(* IEC 61131-3 sources: plc-st-coding-agent/progress/evidence/f14_v3_parallel_20261112/jobs/codex_deepseek-v4pro (part 2) *)

(* ---- public-medium-05.candidate_02.st ---- *)
FUNCTION_BLOCK AutomatedProductionLine
VAR_INPUT
    Mode : BOOL;
    ForwardButton : BOOL;
    ReverseButton : BOOL;
    SensorA : BOOL;
    SensorB : BOOL;
    SensorC : BOOL;
    ButtonA : BOOL;
    ButtonB : BOOL;
    ButtonC : BOOL;
END_VAR
VAR_OUTPUT
    MotorForward : BOOL;
    MotorReverse : BOOL;
    CompletionLight : BOOL;
END_VAR
VAR
    SequenceStep : INT := 0;
END_VAR

MotorForward := FALSE;
MotorReverse := FALSE;
CompletionLight := FALSE;

IF NOT Mode THEN
    MotorForward := ForwardButton AND NOT ReverseButton;
    MotorReverse := ReverseButton AND NOT ForwardButton;
ELSE
    MotorReverse := FALSE;

    CASE SequenceStep OF
        0:
            IF SensorA AND ButtonA THEN
                SequenceStep := 1;
            END_IF;

        1:
            MotorForward := TRUE;
            IF SensorB THEN
                MotorForward := FALSE;
                SequenceStep := 2;
            END_IF;

        2:
            IF ButtonB THEN
                SequenceStep := 3;
            END_IF;

        3:
            MotorForward := TRUE;
            IF SensorC THEN
                MotorForward := FALSE;
                SequenceStep := 4;
            END_IF;

        4:
            IF ButtonC THEN
                SequenceStep := 5;
            END_IF;

        5:
            CompletionLight := SensorC;
            IF NOT SensorC THEN
                CompletionLight := FALSE;
                SequenceStep := 0;
            END_IF;
    END_CASE;
END_IF;

END_FUNCTION_BLOCK

(* ---- public-medium-05.raw_candidate_01.st ---- *)
FUNCTION_BLOCK AutomatedProductionLine
VAR
    SequenceStep : INT := 0;
END_VAR

MotorForward := FALSE;
MotorReverse := FALSE;
CompletionLight := FALSE;

IF NOT Mode THEN
    MotorForward := ForwardButton AND NOT ReverseButton;
    MotorReverse := ReverseButton AND NOT ForwardButton;
    CompletionLight := FALSE;
ELSE
    MotorReverse := FALSE;

    CASE SequenceStep OF
        0:
            IF SensorA AND ButtonA THEN
                SequenceStep := 1;
            END_IF;

        1:
            MotorForward := TRUE;
            IF SensorB THEN
                MotorForward := FALSE;
                SequenceStep := 2;
            END_IF;

        2:
            IF ButtonB THEN
                SequenceStep := 3;
            END_IF;

        3:
            MotorForward := TRUE;
            IF SensorC THEN
                MotorForward := FALSE;
                SequenceStep := 4;
            END_IF;

        4:
            IF ButtonC THEN
                SequenceStep := 5;
            END_IF;

        5:
            CompletionLight := SensorC;
            IF NOT SensorC THEN
                CompletionLight := FALSE;
                SequenceStep := 0;
            END_IF;
    END_CASE;
END_IF;

END_FUNCTION_BLOCK

(* ---- public-medium-05.raw_candidate_02.st ---- *)
FUNCTION_BLOCK AutomatedProductionLine
VAR_INPUT
    Mode : BOOL;
    ForwardButton : BOOL;
    ReverseButton : BOOL;
    SensorA : BOOL;
    SensorB : BOOL;
    SensorC : BOOL;
    ButtonA : BOOL;
    ButtonB : BOOL;
    ButtonC : BOOL;
END_VAR
VAR_OUTPUT
    MotorForward : BOOL;
    MotorReverse : BOOL;
    CompletionLight : BOOL;
END_VAR
VAR
    SequenceStep : INT := 0;
END_VAR

MotorForward := FALSE;
MotorReverse := FALSE;
CompletionLight := FALSE;

IF NOT Mode THEN
    MotorForward := ForwardButton AND NOT ReverseButton;
    MotorReverse := ReverseButton AND NOT ForwardButton;
ELSE
    MotorReverse := FALSE;

    CASE SequenceStep OF
        0:
            IF SensorA AND ButtonA THEN
                SequenceStep := 1;
            END_IF;

        1:
            MotorForward := TRUE;
            IF SensorB THEN
                MotorForward := FALSE;
                SequenceStep := 2;
            END_IF;

        2:
            IF ButtonB THEN
                SequenceStep := 3;
            END_IF;

        3:
            MotorForward := TRUE;
            IF SensorC THEN
                MotorForward := FALSE;
                SequenceStep := 4;
            END_IF;

        4:
            IF ButtonC THEN
                SequenceStep := 5;
            END_IF;

        5:
            CompletionLight := SensorC;
            IF NOT SensorC THEN
                CompletionLight := FALSE;
                SequenceStep := 0;
            END_IF;
    END_CASE;
END_IF;

END_FUNCTION_BLOCK

(* ---- public-medium-06.candidate_01.st ---- *)
FUNCTION_BLOCK SlabThicknessAlarmFaultHistory
VAR_INPUT
    THICKNESS_FAULT : BOOL;
    THICKNESS_SIGNAL_VALID : BOOL;
    CUTTING_RUN : BOOL;
    FaultTimestamp : DINT;
    CycleTime : TIME;
END_VAR
VAR_OUTPUT
    THICKNESS_ALARM : BOOL;
    Slab_Fault_Counter : UINT;
    Slab_Runtime_Accumulator : LTIME;
    Slab_Fault_History : ARRAY[0..4] OF DINT;
END_VAR
VAR
    Initialized : BOOL := FALSE;
    CurrentValidFault : BOOL;
    LastValidFault : BOOL := FALSE;
    AlarmHolding : BOOL := FALSE;
    AlarmHoldTimer : TIME := T#0ms;
    ArrayIndex : INT;
END_VAR

IF NOT Initialized THEN
    THICKNESS_ALARM := FALSE;
    Slab_Fault_Counter := 0;
    Slab_Runtime_Accumulator := TIME_TO_LTIME(T#0ms);
    FOR ArrayIndex := 0 TO 4 DO
        Slab_Fault_History[ArrayIndex] := 0;
    END_FOR;
    AlarmHolding := FALSE;
    AlarmHoldTimer := T#0ms;
    LastValidFault := THICKNESS_SIGNAL_VALID AND THICKNESS_FAULT;
    Initialized := TRUE;
END_IF;

IF NOT THICKNESS_SIGNAL_VALID THEN
    THICKNESS_ALARM := FALSE;
    AlarmHolding := FALSE;
    AlarmHoldTimer := T#0ms;
    LastValidFault := FALSE;
ELSE
    CurrentValidFault := THICKNESS_FAULT;

    IF CurrentValidFault AND NOT LastValidFault THEN
        Slab_Fault_Counter := Slab_Fault_Counter + 1;
        FOR ArrayIndex := 4 TO 1 BY -1 DO
            Slab_Fault_History[ArrayIndex] := Slab_Fault_History[ArrayIndex - 1];
        END_FOR;
        Slab_Fault_History[0] := FaultTimestamp;
    END_IF;

    IF CurrentValidFault THEN
        THICKNESS_ALARM := TRUE;
        AlarmHolding := TRUE;
        AlarmHoldTimer := T#0ms;
    ELSIF AlarmHolding THEN
        AlarmHoldTimer := AlarmHoldTimer + CycleTime;
        THICKNESS_ALARM := TRUE;
        IF AlarmHoldTimer >= T#500ms THEN
            THICKNESS_ALARM := FALSE;
            AlarmHolding := FALSE;
            AlarmHoldTimer := T#0ms;
        END_IF;
    ELSE
        THICKNESS_ALARM := FALSE;
    END_IF;

    LastValidFault := CurrentValidFault;
END_IF;

IF CUTTING_RUN AND THICKNESS_SIGNAL_VALID AND NOT THICKNESS_FAULT THEN
    Slab_Runtime_Accumulator := Slab_Runtime_Accumulator + TIME_TO_LTIME(CycleTime);
END_IF;

END_FUNCTION_BLOCK

(* ---- public-medium-06.candidate_02.st ---- *)
FUNCTION_BLOCK SlabThicknessAlarmFaultHistory
VAR_INPUT
    THICKNESS_FAULT : BOOL;
    THICKNESS_SIGNAL_VALID : BOOL;
    CUTTING_RUN : BOOL;
    FaultTimestamp : DINT;
    CycleTime : TIME;
END_VAR
VAR_OUTPUT
    THICKNESS_ALARM : BOOL;
    Slab_Fault_Counter : UINT;
    Slab_Runtime_Accumulator : LTIME;
    Slab_Fault_History : ARRAY[0..4] OF DINT;
END_VAR
VAR
    PowerUp : BOOL := TRUE;
    LastValidFault : BOOL := FALSE;
    CurrentFault : BOOL;
    AlarmHoldActive : BOOL := FALSE;
    AlarmHoldElapsed : TIME := T#0ms;
    LoopIndex : INT;
END_VAR

IF PowerUp THEN
    THICKNESS_ALARM := FALSE;
    Slab_Fault_Counter := 0;
    Slab_Runtime_Accumulator := TIME_TO_LTIME(T#0ms);
    FOR LoopIndex := 0 TO 4 DO
        Slab_Fault_History[LoopIndex] := 0;
    END_FOR;
    LastValidFault := FALSE;
    AlarmHoldActive := FALSE;
    AlarmHoldElapsed := T#0ms;
    PowerUp := FALSE;
END_IF;

IF NOT THICKNESS_SIGNAL_VALID THEN
    THICKNESS_ALARM := FALSE;
    AlarmHoldActive := FALSE;
    AlarmHoldElapsed := T#0ms;
    LastValidFault := FALSE;
ELSE
    CurrentFault := THICKNESS_FAULT;

    IF CurrentFault AND NOT LastValidFault THEN
        Slab_Fault_Counter := Slab_Fault_Counter + 1;
        FOR LoopIndex := 4 TO 1 BY -1 DO
            Slab_Fault_History[LoopIndex] := Slab_Fault_History[LoopIndex - 1];
        END_FOR;
        Slab_Fault_History[0] := FaultTimestamp;
    END_IF;

    IF CurrentFault THEN
        THICKNESS_ALARM := TRUE;
        AlarmHoldActive := TRUE;
        AlarmHoldElapsed := T#0ms;
    ELSIF AlarmHoldActive THEN
        AlarmHoldElapsed := AlarmHoldElapsed + CycleTime;
        IF AlarmHoldElapsed >= T#500ms THEN
            THICKNESS_ALARM := FALSE;
            AlarmHoldActive := FALSE;
            AlarmHoldElapsed := T#0ms;
        ELSE
            THICKNESS_ALARM := TRUE;
        END_IF;
    ELSE
        THICKNESS_ALARM := FALSE;
    END_IF;

    LastValidFault := CurrentFault;
END_IF;

IF CUTTING_RUN AND THICKNESS_SIGNAL_VALID AND NOT THICKNESS_FAULT THEN
    Slab_Runtime_Accumulator := Slab_Runtime_Accumulator + TIME_TO_LTIME(CycleTime);
END_IF;

END_FUNCTION_BLOCK

(* ---- public-medium-06.raw_candidate_01.st ---- *)
FUNCTION_BLOCK SlabThicknessAlarmFaultHistory
VAR_INPUT
    THICKNESS_FAULT : BOOL;
    THICKNESS_SIGNAL_VALID : BOOL;
    CUTTING_RUN : BOOL;
    FaultTimestamp : DINT;
    CycleTime : TIME;
END_VAR
VAR_OUTPUT
    THICKNESS_ALARM : BOOL;
    Slab_Fault_Counter : UINT;
    Slab_Runtime_Accumulator : LTIME;
    Slab_Fault_History : ARRAY[0..4] OF DINT;
END_VAR
VAR
    Initialized : BOOL := FALSE;
    CurrentValidFault : BOOL;
    LastValidFault : BOOL := FALSE;
    AlarmHolding : BOOL := FALSE;
    AlarmHoldTimer : TIME := T#0ms;
    ArrayIndex : INT;
END_VAR

IF NOT Initialized THEN
    THICKNESS_ALARM := FALSE;
    Slab_Fault_Counter := 0;
    Slab_Runtime_Accumulator := TIME_TO_LTIME(T#0ms);
    FOR ArrayIndex := 0 TO 4 DO
        Slab_Fault_History[ArrayIndex] := 0;
    END_FOR;
    AlarmHolding := FALSE;
    AlarmHoldTimer := T#0ms;
    LastValidFault := THICKNESS_SIGNAL_VALID AND THICKNESS_FAULT;
    Initialized := TRUE;
END_IF;

IF NOT THICKNESS_SIGNAL_VALID THEN
    THICKNESS_ALARM := FALSE;
    AlarmHolding := FALSE;
    AlarmHoldTimer := T#0ms;
    LastValidFault := FALSE;
ELSE
    CurrentValidFault := THICKNESS_FAULT;

    IF CurrentValidFault AND NOT LastValidFault THEN
        Slab_Fault_Counter := Slab_Fault_Counter + 1;
        FOR ArrayIndex := 4 TO 1 BY -1 DO
            Slab_Fault_History[ArrayIndex] := Slab_Fault_History[ArrayIndex - 1];
        END_FOR;
        Slab_Fault_History[0] := FaultTimestamp;
    END_IF;

    IF CurrentValidFault THEN
        THICKNESS_ALARM := TRUE;
        AlarmHolding := TRUE;
        AlarmHoldTimer := T#0ms;
    ELSIF AlarmHolding THEN
        AlarmHoldTimer := AlarmHoldTimer + CycleTime;
        THICKNESS_ALARM := TRUE;
        IF AlarmHoldTimer >= T#500ms THEN
            THICKNESS_ALARM := FALSE;
            AlarmHolding := FALSE;
            AlarmHoldTimer := T#0ms;
        END_IF;
    ELSE
        THICKNESS_ALARM := FALSE;
    END_IF;

    LastValidFault := CurrentValidFault;
END_IF;

IF CUTTING_RUN AND THICKNESS_SIGNAL_VALID AND NOT THICKNESS_FAULT THEN
    Slab_Runtime_Accumulator := Slab_Runtime_Accumulator + TIME_TO_LTIME(CycleTime);
END_IF;

END_FUNCTION_BLOCK

(* ---- public-medium-06.raw_candidate_02.st ---- *)
FUNCTION_BLOCK SlabThicknessAlarmFaultHistory
VAR_INPUT
    THICKNESS_FAULT : BOOL;
    THICKNESS_SIGNAL_VALID : BOOL;
    CUTTING_RUN : BOOL;
    FaultTimestamp : DINT;
    CycleTime : TIME;
END_VAR
VAR_OUTPUT
    THICKNESS_ALARM : BOOL;
    Slab_Fault_Counter : UINT;
    Slab_Runtime_Accumulator : LTIME;
    Slab_Fault_History : ARRAY[0..4] OF DINT;
END_VAR
VAR
    PowerUp : BOOL := TRUE;
    LastValidFault : BOOL := FALSE;
    CurrentFault : BOOL;
    AlarmHoldActive : BOOL := FALSE;
    AlarmHoldElapsed : TIME := T#0ms;
    LoopIndex : INT;
END_VAR

IF PowerUp THEN
    THICKNESS_ALARM := FALSE;
    Slab_Fault_Counter := 0;
    Slab_Runtime_Accumulator := TIME_TO_LTIME(T#0ms);
    FOR LoopIndex := 0 TO 4 DO
        Slab_Fault_History[LoopIndex] := 0;
    END_FOR;
    LastValidFault := FALSE;
    AlarmHoldActive := FALSE;
    AlarmHoldElapsed := T#0ms;
    PowerUp := FALSE;
END_IF;

IF NOT THICKNESS_SIGNAL_VALID THEN
    THICKNESS_ALARM := FALSE;
    AlarmHoldActive := FALSE;
    AlarmHoldElapsed := T#0ms;
    LastValidFault := FALSE;
ELSE
    CurrentFault := THICKNESS_FAULT;

    IF CurrentFault AND NOT LastValidFault THEN
        Slab_Fault_Counter := Slab_Fault_Counter + 1;
        FOR LoopIndex := 4 TO 1 BY -1 DO
            Slab_Fault_History[LoopIndex] := Slab_Fault_History[LoopIndex - 1];
        END_FOR;
        Slab_Fault_History[0] := FaultTimestamp;
    END_IF;

    IF CurrentFault THEN
        THICKNESS_ALARM := TRUE;
        AlarmHoldActive := TRUE;
        AlarmHoldElapsed := T#0ms;
    ELSIF AlarmHoldActive THEN
        AlarmHoldElapsed := AlarmHoldElapsed + CycleTime;
        IF AlarmHoldElapsed >= T#500ms THEN
            THICKNESS_ALARM := FALSE;
            AlarmHoldActive := FALSE;
            AlarmHoldElapsed := T#0ms;
        ELSE
            THICKNESS_ALARM := TRUE;
        END_IF;
    ELSE
        THICKNESS_ALARM := FALSE;
    END_IF;

    LastValidFault := CurrentFault;
END_IF;

IF CUTTING_RUN AND THICKNESS_SIGNAL_VALID AND NOT THICKNESS_FAULT THEN
    Slab_Runtime_Accumulator := Slab_Runtime_Accumulator + TIME_TO_LTIME(CycleTime);
END_IF;

END_FUNCTION_BLOCK

(* ---- public-medium-07.candidate_01.st ---- *)
FUNCTION_BLOCK OfficeHVACMultiModeControl
VAR_INPUT
    OCCUPANCY_DETECTED : BOOL;
    ENERGY_SAVING_MODE : BOOL;
    HVAC_MODE_SELECTOR : INT;
END_VAR
VAR_OUTPUT
    SUPPLY_FAN_RUN : BOOL := FALSE;
    TEMP_SETPOINT_ADJUST : INT := 0;
END_VAR
VAR
    fan_timer : TON;
    setpoint_calc : INT;
END_VAR

fan_timer(IN := OCCUPANCY_DETECTED AND (HVAC_MODE_SELECTOR <> 3), PT := T#30S);
SUPPLY_FAN_RUN := fan_timer.Q;

CASE HVAC_MODE_SELECTOR OF
    0:
        IF OCCUPANCY_DETECTED THEN
            setpoint_calc := 0;
        ELSIF ENERGY_SAVING_MODE THEN
            setpoint_calc := 3;
        ELSE
            setpoint_calc := 2;
        END_IF;
    1:
        IF OCCUPANCY_DETECTED THEN
            setpoint_calc := 0;
        ELSE
            setpoint_calc := 1;
        END_IF;
    2:
        IF OCCUPANCY_DETECTED THEN
            setpoint_calc := 0;
        ELSE
            setpoint_calc := 4;
        END_IF;
    3:
        setpoint_calc := 4;
    ELSE
        setpoint_calc := 0;
END_CASE;

IF setpoint_calc > 4 THEN
    TEMP_SETPOINT_ADJUST := 4;
ELSIF setpoint_calc < -4 THEN
    TEMP_SETPOINT_ADJUST := -4;
ELSE
    TEMP_SETPOINT_ADJUST := setpoint_calc;
END_IF;
END_FUNCTION_BLOCK

(* ---- public-medium-07.raw_candidate_01.st ---- *)
FUNCTION_BLOCK OfficeHVACMultiModeControl
VAR_INPUT
    OCCUPANCY_DETECTED : BOOL;
    ENERGY_SAVING_MODE : BOOL;
    HVAC_MODE_SELECTOR : INT;
END_VAR
VAR_OUTPUT
    SUPPLY_FAN_RUN : BOOL := FALSE;
    TEMP_SETPOINT_ADJUST : INT := 0;
END_VAR
VAR
    fan_timer : TON;
    setpoint_calc : INT;
END_VAR

fan_timer(IN := OCCUPANCY_DETECTED AND (HVAC_MODE_SELECTOR <> 3), PT := T#30S);
SUPPLY_FAN_RUN := fan_timer.Q;

CASE HVAC_MODE_SELECTOR OF
    0:
        IF OCCUPANCY_DETECTED THEN
            setpoint_calc := 0;
        ELSIF ENERGY_SAVING_MODE THEN
            setpoint_calc := 3;
        ELSE
            setpoint_calc := 2;
        END_IF;
    1:
        IF OCCUPANCY_DETECTED THEN
            setpoint_calc := 0;
        ELSE
            setpoint_calc := 1;
        END_IF;
    2:
        IF OCCUPANCY_DETECTED THEN
            setpoint_calc := 0;
        ELSE
            setpoint_calc := 4;
        END_IF;
    3:
        setpoint_calc := 4;
    ELSE
        setpoint_calc := 0;
END_CASE;

IF setpoint_calc > 4 THEN
    TEMP_SETPOINT_ADJUST := 4;
ELSIF setpoint_calc < -4 THEN
    TEMP_SETPOINT_ADJUST := -4;
ELSE
    TEMP_SETPOINT_ADJUST := setpoint_calc;
END_IF;
END_FUNCTION_BLOCK

(* ---- public-medium-08.candidate_01.st ---- *)
FUNCTION_BLOCK IPv4Parser
VAR_INPUT
    ipText : STRING(254);
END_VAR
VAR_OUTPUT
    ipValue : UDINT;
END_VAR
VAR
    bValid : BOOL;
    iPos : INT;
    iLength : INT;
    iCharCode : INT;
    uiCurrentValue : UDINT;
    uiDigitCount : UDINT;
    uiCompletedSegments : UDINT;
    uiAddress : UDINT;
END_VAR

ipValue := 0;
uiAddress := 0;
uiCurrentValue := 0;
uiDigitCount := 0;
uiCompletedSegments := 0;
bValid := TRUE;
iLength := LEN(ipText);

IF (iLength > 0) AND (iLength <= 15) THEN
    FOR iPos := 1 TO iLength BY 1 DO
        iCharCode := BYTE_TO_INT(ipText[iPos]);

        IF (iCharCode >= 48) AND (iCharCode <= 57) THEN
            uiCurrentValue := uiCurrentValue * 10 + INT_TO_UDINT(iCharCode - 48);
            uiDigitCount := uiDigitCount + 1;

            IF uiCurrentValue > 255 THEN
                bValid := FALSE;
                EXIT;
            END_IF;

        ELSIF iCharCode = 46 THEN
            IF (uiDigitCount = 0) OR (uiCompletedSegments >= 3) THEN
                bValid := FALSE;
                EXIT;
            END_IF;

            uiAddress := uiAddress * 256 + uiCurrentValue;
            uiCompletedSegments := uiCompletedSegments + 1;
            uiCurrentValue := 0;
            uiDigitCount := 0;

        ELSE
            bValid := FALSE;
            EXIT;
        END_IF;
    END_FOR;
ELSE
    bValid := FALSE;
END_IF;

IF bValid THEN
    IF (uiDigitCount = 0) OR (uiCompletedSegments <> 3) THEN
        bValid := FALSE;
    ELSE
        uiAddress := uiAddress * 256 + uiCurrentValue;
        ipValue := uiAddress;
    END_IF;
END_IF;

END_FUNCTION_BLOCK

(* ---- public-medium-08.raw_candidate_01.st ---- *)
FUNCTION_BLOCK IPv4Parser
VAR_INPUT
    ipText : STRING(254);
END_VAR
VAR_OUTPUT
    ipValue : UDINT;
END_VAR
VAR
    bValid : BOOL;
    iPos : INT;
    iLength : INT;
    iCharCode : INT;
    uiCurrentValue : UDINT;
    uiDigitCount : UDINT;
    uiCompletedSegments : UDINT;
    uiAddress : UDINT;
END_VAR

ipValue := 0;
uiAddress := 0;
uiCurrentValue := 0;
uiDigitCount := 0;
uiCompletedSegments := 0;
bValid := TRUE;
iLength := LEN(ipText);

IF (iLength > 0) AND (iLength <= 15) THEN
    FOR iPos := 1 TO iLength BY 1 DO
        iCharCode := BYTE_TO_INT(ipText[iPos]);

        IF (iCharCode >= 48) AND (iCharCode <= 57) THEN
            uiCurrentValue := uiCurrentValue * 10 + INT_TO_UDINT(iCharCode - 48);
            uiDigitCount := uiDigitCount + 1;

            IF uiCurrentValue > 255 THEN
                bValid := FALSE;
                EXIT;
            END_IF;

        ELSIF iCharCode = 46 THEN
            IF (uiDigitCount = 0) OR (uiCompletedSegments >= 3) THEN
                bValid := FALSE;
                EXIT;
            END_IF;

            uiAddress := uiAddress * 256 + uiCurrentValue;
            uiCompletedSegments := uiCompletedSegments + 1;
            uiCurrentValue := 0;
            uiDigitCount := 0;

        ELSE
            bValid := FALSE;
            EXIT;
        END_IF;
    END_FOR;
ELSE
    bValid := FALSE;
END_IF;

IF bValid THEN
    IF (uiDigitCount = 0) OR (uiCompletedSegments <> 3) THEN
        bValid := FALSE;
    ELSE
        uiAddress := uiAddress * 256 + uiCurrentValue;
        ipValue := uiAddress;
    END_IF;
END_IF;

END_FUNCTION_BLOCK

(* ---- self-easy-01.candidate_01.st ---- *)
FUNCTION_BLOCK FB
VAR_INPUT
    enable : BOOL;
    values : ARRAY[1..8] OF INT;
    count : INT;
    avgEnable : BOOL;
END_VAR
VAR_OUTPUT
    avgOut : REAL;
END_VAR
VAR
    sampleCount : INT;
    total : LINT;
    idx : INT;
END_VAR

IF enable AND avgEnable AND (count > 0) THEN
    IF count > 8 THEN
        sampleCount := 8;
    ELSE
        sampleCount := count;
    END_IF;

    total := LINT#0;

    FOR idx := 1 TO sampleCount BY 1 DO
        total := total + INT_TO_LINT(values[idx]);
    END_FOR;

    avgOut := LINT_TO_REAL(total) / INT_TO_REAL(sampleCount);
END_IF;

END_FUNCTION_BLOCK

(* ---- self-easy-01.raw_candidate_01.st ---- *)
FUNCTION_BLOCK FB
VAR_INPUT
    enable : BOOL;
    values : ARRAY[1..8] OF INT;
    count : INT;
    avgEnable : BOOL;
END_VAR
VAR_OUTPUT
    avgOut : REAL;
END_VAR
VAR
    sampleCount : INT;
    total : LINT;
    idx : INT;
END_VAR

IF enable AND avgEnable AND (count > 0) THEN
    IF count > 8 THEN
        sampleCount := 8;
    ELSE
        sampleCount := count;
    END_IF;

    total := LINT#0;

    FOR idx := 1 TO sampleCount BY 1 DO
        total := total + INT_TO_LINT(values[idx]);
    END_FOR;

    avgOut := LINT_TO_REAL(total) / INT_TO_REAL(sampleCount);
END_IF;

END_FUNCTION_BLOCK

(* ---- self-easy-02.candidate_01.st ---- *)
FUNCTION_BLOCK FB
VAR_INPUT
    tankLevel : REAL;
    outletFlow : REAL;
    inletPermit : BOOL;
    resetBtn : BOOL;
END_VAR
VAR_OUTPUT
    pumpRun : BOOL;
    alarmHigh : BOOL;
    alarmLow : BOOL;
    outletValveOpen : BOOL;
END_VAR
VAR
    highLatched : BOOL := FALSE;
    lowLatched : BOOL := FALSE;
    prevReset : BOOL := FALSE;
    resetRising : BOOL;
    oldHigh : BOOL;
    oldLow : BOOL;
END_VAR

resetRising := resetBtn AND NOT prevReset;

oldHigh := highLatched;
oldLow := lowLatched;

highLatched := (tankLevel >= 85.0) OR (oldHigh AND NOT resetRising);
lowLatched := (tankLevel <= 15.0) OR (oldLow AND NOT resetRising);

alarmHigh := highLatched;
alarmLow := lowLatched;

pumpRun := inletPermit AND NOT alarmHigh AND NOT alarmLow;
outletValveOpen := NOT alarmLow;

prevReset := resetBtn;
END_FUNCTION_BLOCK

(* ---- self-easy-02.raw_candidate_01.st ---- *)
FUNCTION_BLOCK FB
VAR_INPUT
    tankLevel : REAL;
    outletFlow : REAL;
    inletPermit : BOOL;
    resetBtn : BOOL;
END_VAR
VAR_OUTPUT
    pumpRun : BOOL;
    alarmHigh : BOOL;
    alarmLow : BOOL;
    outletValveOpen : BOOL;
END_VAR
VAR
    highLatched : BOOL := FALSE;
    lowLatched : BOOL := FALSE;
    prevReset : BOOL := FALSE;
    resetRising : BOOL;
    oldHigh : BOOL;
    oldLow : BOOL;
END_VAR

resetRising := resetBtn AND NOT prevReset;

oldHigh := highLatched;
oldLow := lowLatched;

highLatched := (tankLevel >= 85.0) OR (oldHigh AND NOT resetRising);
lowLatched := (tankLevel <= 15.0) OR (oldLow AND NOT resetRising);

alarmHigh := highLatched;
alarmLow := lowLatched;

pumpRun := inletPermit AND NOT alarmHigh AND NOT alarmLow;
outletValveOpen := NOT alarmLow;

prevReset := resetBtn;
END_FUNCTION_BLOCK

(* ---- self-hard-01.candidate_01.st ---- *)
FUNCTION_BLOCK FB
VAR_INPUT
    flowLow : BOOL;
    ackBtn : BOOL;
    sensorOK : BOOL;
END_VAR
VAR_OUTPUT
    alarmActive : BOOL;
    alarmAcked : BOOL;
    highHigh : BOOL;
END_VAR
VAR
    prevAck : BOOL;
    prevFlowLow : BOOL;
    prevAlarmActive : BOOL;
    prevAlarmAcked : BOOL;
    ackRise : BOOL;
END_VAR

ackRise := ackBtn AND NOT prevAck;

highHigh := NOT sensorOK;

alarmActive := flowLow OR (prevAlarmActive AND NOT ackRise AND NOT (prevFlowLow AND prevAlarmAcked));

alarmAcked := alarmActive AND (NOT flowLow OR ackRise OR (prevFlowLow AND prevAlarmActive AND prevAlarmAcked));

prevAck := ackBtn;
prevFlowLow := flowLow;
prevAlarmActive := alarmActive;
prevAlarmAcked := alarmAcked;

END_FUNCTION_BLOCK

(* ---- self-hard-01.raw_candidate_01.st ---- *)
FUNCTION_BLOCK FB
VAR_INPUT
    flowLow : BOOL;
    ackBtn : BOOL;
    sensorOK : BOOL;
END_VAR
VAR_OUTPUT
    alarmActive : BOOL;
    alarmAcked : BOOL;
    highHigh : BOOL;
END_VAR
VAR
    prevAck : BOOL;
    prevFlowLow : BOOL;
    prevAlarmActive : BOOL;
    prevAlarmAcked : BOOL;
    ackRise : BOOL;
END_VAR

ackRise := ackBtn AND NOT prevAck;

highHigh := NOT sensorOK;

alarmActive := flowLow OR (prevAlarmActive AND NOT ackRise AND NOT (prevFlowLow AND prevAlarmAcked));

alarmAcked := alarmActive AND (NOT flowLow OR ackRise OR (prevFlowLow AND prevAlarmActive AND prevAlarmAcked));

prevAck := ackBtn;
prevFlowLow := flowLow;
prevAlarmActive := alarmActive;
prevAlarmAcked := alarmAcked;

END_FUNCTION_BLOCK

(* ---- self-hard-02.candidate_01.st ---- *)
FUNCTION_BLOCK FB
VAR_INPUT
    startBtn    : BOOL;
    abortBtn    : BOOL;
    setpoint    : REAL;
    pv          : REAL;
    maxDuration : INT;
END_VAR
VAR_OUTPUT
    elapsed : INT;
    phase   : INT;
    timeout : BOOL;
END_VAR
VAR
    prevStart    : BOOL;
    statePhase   : INT;
    stateElapsed : INT;
    stateTimeout : BOOL;
END_VAR

IF abortBtn THEN
    statePhase := 9;
ELSIF startBtn AND NOT prevStart THEN
    statePhase   := 1;
    stateElapsed := 0;
    stateTimeout := FALSE;
ELSE
    IF statePhase = 1 OR statePhase = 2 THEN
        stateElapsed := stateElapsed + 1;
        IF stateElapsed >= maxDuration THEN
            stateTimeout := TRUE;
            statePhase   := 3;
        ELSIF statePhase = 2 THEN
            stateTimeout := FALSE;
            statePhase   := 2;
        ELSIF pv >= setpoint THEN
            stateTimeout := FALSE;
            statePhase   := 2;
        ELSE
            stateTimeout := FALSE;
            statePhase   := 1;
        END_IF;
    END_IF;
END_IF;

phase   := statePhase;
elapsed := stateElapsed;
timeout := stateTimeout;

prevStart := startBtn;

END_FUNCTION_BLOCK

(* ---- self-hard-02.raw_candidate_01.st ---- *)
FUNCTION_BLOCK FB
VAR_INPUT
    startBtn    : BOOL;
    abortBtn    : BOOL;
    setpoint    : REAL;
    pv          : REAL;
    maxDuration : INT;
END_VAR
VAR_OUTPUT
    elapsed : INT;
    phase   : INT;
    timeout : BOOL;
END_VAR
VAR
    prevStart    : BOOL;
    statePhase   : INT;
    stateElapsed : INT;
    stateTimeout : BOOL;
END_VAR

IF abortBtn THEN
    statePhase := 9;
ELSIF startBtn AND NOT prevStart THEN
    statePhase   := 1;
    stateElapsed := 0;
    stateTimeout := FALSE;
ELSE
    IF statePhase = 1 OR statePhase = 2 THEN
        stateElapsed := stateElapsed + 1;
        IF stateElapsed >= maxDuration THEN
            stateTimeout := TRUE;
            statePhase   := 3;
        ELSIF statePhase = 2 THEN
            stateTimeout := FALSE;
            statePhase   := 2;
        ELSIF pv >= setpoint THEN
            stateTimeout := FALSE;
            statePhase   := 2;
        ELSE
            stateTimeout := FALSE;
            statePhase   := 1;
        END_IF;
    END_IF;
END_IF;

phase   := statePhase;
elapsed := stateElapsed;
timeout := stateTimeout;

prevStart := startBtn;

END_FUNCTION_BLOCK

(* ---- self-hard-03.candidate_01.st ---- *)
FUNCTION_BLOCK FB
VAR
    qcnt : INT := 0;
    pushPrev : BOOL := FALSE;
    popPrev : BOOL := FALSE;
    pushRise : BOOL;
    popRise : BOOL;
    idx : INT;
END_VAR

pushRise := pushEn AND NOT pushPrev;
popRise := popEn AND NOT popPrev;

IF popRise AND qcnt > 0 THEN
    FOR idx := 1 TO qcnt - 1 DO
        fifo[idx] := fifo[idx + 1];
    END_FOR;
    qcnt := qcnt - 1;
END_IF;

IF pushRise AND qcnt < 8 THEN
    fifo[qcnt + 1] := pushItem;
    qcnt := qcnt + 1;
END_IF;

count := qcnt;
full := (qcnt = 8);
empty := (qcnt = 0);

IF qcnt = 0 THEN
    head := 0;
ELSE
    head := fifo[1];
END_IF;

pushPrev := pushEn;
popPrev := popEn;
END_FUNCTION_BLOCK

(* ---- self-hard-03.candidate_02.st ---- *)
FUNCTION_BLOCK FB
VAR_INPUT
    pushEn : BOOL;
    pushItem : INT;
    popEn : BOOL;
END_VAR
VAR_IN_OUT
    fifo : ARRAY[1..8] OF INT;
END_VAR
VAR_OUTPUT
    count : INT;
    full : BOOL;
    empty : BOOL;
    head : INT;
END_VAR
VAR
    qcnt : INT := 0;
    pushPrev : BOOL := FALSE;
    popPrev : BOOL := FALSE;
    pushRise : BOOL;
    popRise : BOOL;
    idx : INT;
END_VAR

pushRise := pushEn AND NOT pushPrev;
popRise := popEn AND NOT popPrev;

IF popRise AND qcnt > 0 THEN
    FOR idx := 1 TO qcnt - 1 DO
        fifo[idx] := fifo[idx + 1];
    END_FOR;
    qcnt := qcnt - 1;
END_IF;

IF pushRise AND qcnt < 8 THEN
    fifo[qcnt + 1] := pushItem;
    qcnt := qcnt + 1;
END_IF;

count := qcnt;
full := (qcnt = 8);
empty := (qcnt = 0);

IF qcnt = 0 THEN
    head := 0;
ELSE
    head := fifo[1];
END_IF;

pushPrev := pushEn;
popPrev := popEn;
END_FUNCTION_BLOCK

(* ---- self-hard-03.raw_candidate_01.st ---- *)
FUNCTION_BLOCK FB
VAR
    qcnt : INT := 0;
    pushPrev : BOOL := FALSE;
    popPrev : BOOL := FALSE;
    pushRise : BOOL;
    popRise : BOOL;
    idx : INT;
END_VAR

pushRise := pushEn AND NOT pushPrev;
popRise := popEn AND NOT popPrev;

IF popRise AND qcnt > 0 THEN
    FOR idx := 1 TO qcnt - 1 DO
        fifo[idx] := fifo[idx + 1];
    END_FOR;
    qcnt := qcnt - 1;
END_IF;

IF pushRise AND qcnt < 8 THEN
    fifo[qcnt + 1] := pushItem;
    qcnt := qcnt + 1;
END_IF;

count := qcnt;
full := (qcnt = 8);
empty := (qcnt = 0);

IF qcnt = 0 THEN
    head := 0;
ELSE
    head := fifo[1];
END_IF;

pushPrev := pushEn;
popPrev := popEn;
END_FUNCTION_BLOCK

(* ---- self-hard-03.raw_candidate_02.st ---- *)
FUNCTION_BLOCK FB
VAR_INPUT
    pushEn : BOOL;
    pushItem : INT;
    popEn : BOOL;
END_VAR
VAR_IN_OUT
    fifo : ARRAY[1..8] OF INT;
END_VAR
VAR_OUTPUT
    count : INT;
    full : BOOL;
    empty : BOOL;
    head : INT;
END_VAR
VAR
    qcnt : INT := 0;
    pushPrev : BOOL := FALSE;
    popPrev : BOOL := FALSE;
    pushRise : BOOL;
    popRise : BOOL;
    idx : INT;
END_VAR

pushRise := pushEn AND NOT pushPrev;
popRise := popEn AND NOT popPrev;

IF popRise AND qcnt > 0 THEN
    FOR idx := 1 TO qcnt - 1 DO
        fifo[idx] := fifo[idx + 1];
    END_FOR;
    qcnt := qcnt - 1;
END_IF;

IF pushRise AND qcnt < 8 THEN
    fifo[qcnt + 1] := pushItem;
    qcnt := qcnt + 1;
END_IF;

count := qcnt;
full := (qcnt = 8);
empty := (qcnt = 0);

IF qcnt = 0 THEN
    head := 0;
ELSE
    head := fifo[1];
END_IF;

pushPrev := pushEn;
popPrev := popEn;
END_FUNCTION_BLOCK

(* ---- self-hard-04.candidate_01.st ---- *)
FUNCTION_BLOCK FB
VAR_INPUT
    demand : INT;
    runHours : ARRAY[1..5] OF LINT;
    rotated : BOOL;
END_VAR
VAR_OUTPUT
    leadPump : INT;
    lagPump : INT;
    runningCount : INT;
END_VAR
VAR
    demandClipped : INT;
    prevLeadPump : INT := 0;
    prevLagPump : INT := 0;
    prevRunningCount : INT := 0;
    minPump : INT;
    minHours : LINT;
    bestLagPump : INT;
    bestLagHours : LINT;
    idx : INT;
    leadChanged : BOOL;
    countRose : BOOL;
    rotationThreshold : LINT := 50;
END_VAR

demandClipped := demand;
IF demandClipped < 0 THEN
    demandClipped := 0;
ELSIF demandClipped > 5 THEN
    demandClipped := 5;
END_IF;

runningCount := demandClipped;

IF demandClipped <= 0 THEN
    leadPump := 0;
    lagPump := 0;
ELSE
    minPump := 1;
    minHours := runHours[1];
    FOR idx := 2 TO 5 BY 1 DO
        IF runHours[idx] < minHours THEN
            minPump := idx;
            minHours := runHours[idx];
        END_IF;
    END_FOR;

    IF prevLeadPump = 0 THEN
        leadPump := minPump;
    ELSIF rotated THEN
        IF runHours[prevLeadPump] - minHours > rotationThreshold THEN
            leadPump := minPump;
        ELSE
            leadPump := prevLeadPump;
        END_IF;
    ELSE
        leadPump := prevLeadPump;
    END_IF;

    IF demandClipped < 2 THEN
        lagPump := 0;
    ELSE
        leadChanged := leadPump <> prevLeadPump;
        countRose := demandClipped > prevRunningCount;

        IF leadChanged OR countRose THEN
            bestLagPump := 0;
            FOR idx := 1 TO 5 BY 1 DO
                IF idx <> leadPump THEN
                    IF bestLagPump = 0 THEN
                        bestLagPump := idx;
                        bestLagHours := runHours[idx];
                    ELSIF runHours[idx] < bestLagHours THEN
                        bestLagPump := idx;
                        bestLagHours := runHours[idx];
                    END_IF;
                END_IF;
            END_FOR;
            lagPump := bestLagPump;
        ELSE
            lagPump := prevLagPump;
        END_IF;
    END_IF;
END_IF;

prevLeadPump := leadPump;
prevLagPump := lagPump;
prevRunningCount := runningCount;

END_FUNCTION_BLOCK

(* ---- self-hard-04.raw_candidate_01.st ---- *)
FUNCTION_BLOCK FB
VAR_INPUT
    demand : INT;
    runHours : ARRAY[1..5] OF LINT;
    rotated : BOOL;
END_VAR
VAR_OUTPUT
    leadPump : INT;
    lagPump : INT;
    runningCount : INT;
END_VAR
VAR
    demandClipped : INT;
    prevLeadPump : INT := 0;
    prevLagPump : INT := 0;
    prevRunningCount : INT := 0;
    minPump : INT;
    minHours : LINT;
    bestLagPump : INT;
    bestLagHours : LINT;
    idx : INT;
    leadChanged : BOOL;
    countRose : BOOL;
    rotationThreshold : LINT := 50;
END_VAR

demandClipped := demand;
IF demandClipped < 0 THEN
    demandClipped := 0;
ELSIF demandClipped > 5 THEN
    demandClipped := 5;
END_IF;

runningCount := demandClipped;

IF demandClipped <= 0 THEN
    leadPump := 0;
    lagPump := 0;
ELSE
    minPump := 1;
    minHours := runHours[1];
    FOR idx := 2 TO 5 BY 1 DO
        IF runHours[idx] < minHours THEN
            minPump := idx;
            minHours := runHours[idx];
        END_IF;
    END_FOR;

    IF prevLeadPump = 0 THEN
        leadPump := minPump;
    ELSIF rotated THEN
        IF runHours[prevLeadPump] - minHours > rotationThreshold THEN
            leadPump := minPump;
        ELSE
            leadPump := prevLeadPump;
        END_IF;
    ELSE
        leadPump := prevLeadPump;
    END_IF;

    IF demandClipped < 2 THEN
        lagPump := 0;
    ELSE
        leadChanged := leadPump <> prevLeadPump;
        countRose := demandClipped > prevRunningCount;

        IF leadChanged OR countRose THEN
            bestLagPump := 0;
            FOR idx := 1 TO 5 BY 1 DO
                IF idx <> leadPump THEN
                    IF bestLagPump = 0 THEN
                        bestLagPump := idx;
                        bestLagHours := runHours[idx];
                    ELSIF runHours[idx] < bestLagHours THEN
                        bestLagPump := idx;
                        bestLagHours := runHours[idx];
                    END_IF;
                END_IF;
            END_FOR;
            lagPump := bestLagPump;
        ELSE
            lagPump := prevLagPump;
        END_IF;
    END_IF;
END_IF;

prevLeadPump := leadPump;
prevLagPump := lagPump;
prevRunningCount := runningCount;

END_FUNCTION_BLOCK

(* ---- self-hard-05.candidate_01.st ---- *)
FUNCTION_BLOCK FB
VAR_INPUT
    runRequest : BOOL;
    flameOK : BOOL;
    o2Valid : BOOL;
    o2PV : REAL;
    baseAir : REAL;
    resetBtn : BOOL;
END_VAR
VAR_OUTPUT
    fuelPermit : BOOL;
    trimEnable : BOOL;
    airTrim : REAL;
    airCommand : REAL;
    tripLatched : BOOL;
    o2Fault : BOOL;
END_VAR
VAR
    prevReset : BOOL;
    prevTrip : BOOL;
    resetRise : BOOL;
    rawTrim : REAL;
    rawCmd : REAL;
END_VAR

resetRise := resetBtn AND NOT prevReset;

tripLatched := (runRequest AND NOT flameOK)
    OR (prevTrip AND NOT (resetRise AND NOT runRequest AND NOT flameOK));

fuelPermit := runRequest AND flameOK AND NOT tripLatched;

o2Fault := NOT o2Valid OR o2PV < 0.0 OR o2PV > 21.0;

trimEnable := fuelPermit AND NOT o2Fault;

IF trimEnable THEN
    rawTrim := 2.0 * (2.0 - o2PV);
    IF rawTrim < -10.0 THEN
        airTrim := -10.0;
    ELSIF rawTrim > 10.0 THEN
        airTrim := 10.0;
    ELSE
        airTrim := rawTrim;
    END_IF;
ELSE
    airTrim := 0.0;
END_IF;

IF NOT fuelPermit THEN
    airCommand := 0.0;
ELSE
    rawCmd := baseAir + airTrim;
    IF rawCmd < 0.0 THEN
        airCommand := 0.0;
    ELSIF rawCmd > 100.0 THEN
        airCommand := 100.0;
    ELSE
        airCommand := rawCmd;
    END_IF;
END_IF;

prevReset := resetBtn;
prevTrip := tripLatched;

END_FUNCTION_BLOCK

(* ---- self-hard-05.raw_candidate_01.st ---- *)
FUNCTION_BLOCK FB
VAR_INPUT
    runRequest : BOOL;
    flameOK : BOOL;
    o2Valid : BOOL;
    o2PV : REAL;
    baseAir : REAL;
    resetBtn : BOOL;
END_VAR
VAR_OUTPUT
    fuelPermit : BOOL;
    trimEnable : BOOL;
    airTrim : REAL;
    airCommand : REAL;
    tripLatched : BOOL;
    o2Fault : BOOL;
END_VAR
VAR
    prevReset : BOOL;
    prevTrip : BOOL;
    resetRise : BOOL;
    rawTrim : REAL;
    rawCmd : REAL;
END_VAR

resetRise := resetBtn AND NOT prevReset;

tripLatched := (runRequest AND NOT flameOK)
    OR (prevTrip AND NOT (resetRise AND NOT runRequest AND NOT flameOK));

fuelPermit := runRequest AND flameOK AND NOT tripLatched;

o2Fault := NOT o2Valid OR o2PV < 0.0 OR o2PV > 21.0;

trimEnable := fuelPermit AND NOT o2Fault;

IF trimEnable THEN
    rawTrim := 2.0 * (2.0 - o2PV);
    IF rawTrim < -10.0 THEN
        airTrim := -10.0;
    ELSIF rawTrim > 10.0 THEN
        airTrim := 10.0;
    ELSE
        airTrim := rawTrim;
    END_IF;
ELSE
    airTrim := 0.0;
END_IF;

IF NOT fuelPermit THEN
    airCommand := 0.0;
ELSE
    rawCmd := baseAir + airTrim;
    IF rawCmd < 0.0 THEN
        airCommand := 0.0;
    ELSIF rawCmd > 100.0 THEN
        airCommand := 100.0;
    ELSE
        airCommand := rawCmd;
    END_IF;
END_IF;

prevReset := resetBtn;
prevTrip := tripLatched;

END_FUNCTION_BLOCK

(* ---- self-hard-06.candidate_01.st ---- *)
FUNCTION_BLOCK FB
VAR_INPUT
    runRequest : BOOL;
    pressure : REAL;
    pressureValid : BOOL;
    fuelFlow : REAL;
    steamFlow : REAL;
    outletCmd : INT;
    outletFeedback : INT;
    resetBtn : BOOL;
END_VAR
VAR_OUTPUT
    tripLatched : BOOL;
    fuelPermit : BOOL;
    currentCauseMask : WORD;
    latchedCauseMask : WORD;
    diagnosticActive : BOOL;
END_VAR
VAR
    prevReset : BOOL;
    prevTrip : BOOL;
    valveCnt : INT;
    tripNow : BOOL;
    validOverpressure : BOOL;
    valveJamCondition : BOOL;
    burnCondition : BOOL;
    valveJamBit : BOOL;
    burnBit : BOOL;
    resetEdge : BOOL;
    legalReset : BOOL;
    nextTrip : BOOL;
    currentMask : WORD;
    latchedStore : WORD;
END_VAR

resetEdge := resetBtn AND NOT prevReset;
legalReset := resetEdge AND NOT runRequest AND pressureValid AND (pressure <= 4200.0);
validOverpressure := runRequest AND pressureValid AND (pressure >= 4500.0);
valveJamCondition := validOverpressure AND (outletCmd >= 50) AND (outletFeedback <= 10);
burnCondition := validOverpressure AND (fuelFlow >= 4.0) AND (steamFlow <= 10.0);

IF valveJamCondition THEN
    IF valveCnt < 3 THEN
        valveCnt := valveCnt + 1;
    END_IF;
ELSE
    valveCnt := 0;
END_IF;

valveJamBit := valveCnt >= 3;
burnBit := burnCondition;

IF runRequest AND NOT pressureValid THEN
    currentMask := WORD#16#0001;
ELSIF validOverpressure THEN
    IF valveJamBit AND burnBit THEN
        currentMask := WORD#16#0006;
    ELSIF valveJamBit THEN
        currentMask := WORD#16#0002;
    ELSIF burnBit THEN
        currentMask := WORD#16#0004;
    ELSE
        currentMask := WORD#16#0008;
    END_IF;
ELSE
    currentMask := WORD#16#0000;
END_IF;

tripNow := runRequest AND (NOT pressureValid OR (pressure >= 4500.0));
IF tripNow THEN
    nextTrip := TRUE;
ELSIF legalReset THEN
    nextTrip := FALSE;
ELSE
    nextTrip := prevTrip;
END_IF;

IF nextTrip THEN
    latchedStore := latchedStore OR currentMask;
ELSE
    latchedStore := WORD#16#0000;
END_IF;

tripLatched := nextTrip;
fuelPermit := runRequest AND NOT nextTrip;
currentCauseMask := currentMask;
latchedCauseMask := latchedStore;
diagnosticActive := currentMask <> WORD#16#0000;

prevReset := resetBtn;
prevTrip := nextTrip;
END_FUNCTION_BLOCK

(* ---- self-hard-06.raw_candidate_01.st ---- *)
FUNCTION_BLOCK FB
VAR_INPUT
    runRequest : BOOL;
    pressure : REAL;
    pressureValid : BOOL;
    fuelFlow : REAL;
    steamFlow : REAL;
    outletCmd : INT;
    outletFeedback : INT;
    resetBtn : BOOL;
END_VAR
VAR_OUTPUT
    tripLatched : BOOL;
    fuelPermit : BOOL;
    currentCauseMask : WORD;
    latchedCauseMask : WORD;
    diagnosticActive : BOOL;
END_VAR
VAR
    prevReset : BOOL;
    prevTrip : BOOL;
    valveCnt : INT;
    tripNow : BOOL;
    validOverpressure : BOOL;
    valveJamCondition : BOOL;
    burnCondition : BOOL;
    valveJamBit : BOOL;
    burnBit : BOOL;
    resetEdge : BOOL;
    legalReset : BOOL;
    nextTrip : BOOL;
    currentMask : WORD;
    latchedStore : WORD;
END_VAR

resetEdge := resetBtn AND NOT prevReset;
legalReset := resetEdge AND NOT runRequest AND pressureValid AND (pressure <= 4200.0);
validOverpressure := runRequest AND pressureValid AND (pressure >= 4500.0);
valveJamCondition := validOverpressure AND (outletCmd >= 50) AND (outletFeedback <= 10);
burnCondition := validOverpressure AND (fuelFlow >= 4.0) AND (steamFlow <= 10.0);

IF valveJamCondition THEN
    IF valveCnt < 3 THEN
        valveCnt := valveCnt + 1;
    END_IF;
ELSE
    valveCnt := 0;
END_IF;

valveJamBit := valveCnt >= 3;
burnBit := burnCondition;

IF runRequest AND NOT pressureValid THEN
    currentMask := WORD#16#0001;
ELSIF validOverpressure THEN
    IF valveJamBit AND burnBit THEN
        currentMask := WORD#16#0006;
    ELSIF valveJamBit THEN
        currentMask := WORD#16#0002;
    ELSIF burnBit THEN
        currentMask := WORD#16#0004;
    ELSE
        currentMask := WORD#16#0008;
    END_IF;
ELSE
    currentMask := WORD#16#0000;
END_IF;

tripNow := runRequest AND (NOT pressureValid OR (pressure >= 4500.0));
IF tripNow THEN
    nextTrip := TRUE;
ELSIF legalReset THEN
    nextTrip := FALSE;
ELSE
    nextTrip := prevTrip;
END_IF;

IF nextTrip THEN
    latchedStore := latchedStore OR currentMask;
ELSE
    latchedStore := WORD#16#0000;
END_IF;

tripLatched := nextTrip;
fuelPermit := runRequest AND NOT nextTrip;
currentCauseMask := currentMask;
latchedCauseMask := latchedStore;
diagnosticActive := currentMask <> WORD#16#0000;

prevReset := resetBtn;
prevTrip := nextTrip;
END_FUNCTION_BLOCK

(* ---- self-hard-07.candidate_01.st ---- *)
FUNCTION_BLOCK FB
VAR_INPUT
    mode : INT;
    resetBtn : BOOL;
    scanSeconds : REAL;
    tempSP : REAL;
    tempPV : REAL;
    flowPV : REAL;
    manualFlowSP : REAL;
    manualValve : REAL;
END_VAR
VAR_OUTPUT
    flowSP : REAL;
    valveCommand : REAL;
    fault : BOOL;
    normalMode : BOOL;
END_VAR
VAR
    initDone : BOOL := FALSE;
    prevMode : INT := 0;
    prevReset : BOOL := FALSE;
    prevFlowSP : REAL := 0.0;
    prevValveCommand : REAL := 0.0;
    accT : REAL := 0.0;
    accF : REAL := 0.0;
    tempError : REAL;
    flowError : REAL;
    trialT : REAL;
    trialF : REAL;
    rawFlow : REAL;
    rawValve : REAL;
    modeChanged : BOOL;
    resetRise : BOOL;
END_VAR

fault := (mode < 0) OR (mode > 2) OR (scanSeconds <= 0.0) OR (scanSeconds > 10.0);
resetRise := resetBtn AND NOT prevReset;
normalMode := FALSE;

IF NOT initDone THEN
    flowSP := manualFlowSP;
    valveCommand := manualValve;
    tempError := tempSP - tempPV;
    accT := flowSP - 1.0 * tempError;
    flowError := flowSP - flowPV;
    accF := valveCommand - 2.0 * flowError;
ELSE
    modeChanged := mode <> prevMode;

    IF resetRise THEN
        flowSP := manualFlowSP;
        valveCommand := manualValve;
        tempError := tempSP - tempPV;
        accT := flowSP - 1.0 * tempError;
        flowError := flowSP - flowPV;
        accF := valveCommand - 2.0 * flowError;
    ELSIF fault THEN
        flowSP := manualFlowSP;
        valveCommand := manualValve;
        tempError := tempSP - tempPV;
        accT := flowSP - 1.0 * tempError;
        flowError := flowSP - flowPV;
        accF := valveCommand - 2.0 * flowError;
    ELSIF modeChanged THEN
        IF mode = 2 THEN
            flowSP := prevFlowSP;
            valveCommand := prevValveCommand;
            tempError := tempSP - tempPV;
            accT := flowSP - 1.0 * tempError;
            flowError := flowSP - flowPV;
            accF := valveCommand - 2.0 * flowError;
        ELSE
            flowSP := manualFlowSP;
            valveCommand := prevValveCommand;
            tempError := tempSP - tempPV;
            accT := flowSP - 1.0 * tempError;
            flowError := flowSP - flowPV;
            accF := valveCommand - 2.0 * flowError;
        END_IF;
    ELSE
        normalMode := TRUE;
        IF mode = 0 THEN
            flowSP := manualFlowSP;
            valveCommand := manualValve;
            tempError := tempSP - tempPV;
            accT := flowSP - 1.0 * tempError;
            flowError := flowSP - flowPV;
            accF := valveCommand - 2.0 * flowError;
        ELSIF mode = 1 THEN
            flowSP := manualFlowSP;
            flowError := flowSP - flowPV;
            trialF := accF + 0.5 * flowError * scanSeconds;
            rawValve := 2.0 * flowError + trialF;
            IF rawValve < 0.0 THEN
                valveCommand := 0.0;
            ELSIF rawValve > 100.0 THEN
                valveCommand := 100.0;
            ELSE
                valveCommand := rawValve;
            END_IF;
            accF := valveCommand - 2.0 * flowError;
            tempError := tempSP - tempPV;
            accT := flowSP - 1.0 * tempError;
        ELSE
            tempError := tempSP - tempPV;
            trialT := accT + 0.2 * tempError * scanSeconds;
            rawFlow := 1.0 * tempError + trialT;
            IF rawFlow < 0.0 THEN
                flowSP := 0.0;
            ELSIF rawFlow > 50.0 THEN
                flowSP := 50.0;
            ELSE
                flowSP := rawFlow;
            END_IF;
            accT := flowSP - 1.0 * tempError;

            flowError := flowSP - flowPV;
            trialF := accF + 0.5 * flowError * scanSeconds;
            rawValve := 2.0 * flowError + trialF;
            IF rawValve < 0.0 THEN
                valveCommand := 0.0;
            ELSIF rawValve > 100.0 THEN
                valveCommand := 100.0;
            ELSE
                valveCommand := rawValve;
            END_IF;
            accF := valveCommand - 2.0 * flowError;
        END_IF;
    END_IF;
END_IF;

prevMode := mode;
prevReset := resetBtn;
prevFlowSP := flowSP;
prevValveCommand := valveCommand;
initDone := TRUE;
END_FUNCTION_BLOCK

(* ---- self-hard-07.raw_candidate_01.st ---- *)
FUNCTION_BLOCK FB
VAR_INPUT
    mode : INT;
    resetBtn : BOOL;
    scanSeconds : REAL;
    tempSP : REAL;
    tempPV : REAL;
    flowPV : REAL;
    manualFlowSP : REAL;
    manualValve : REAL;
END_VAR
VAR_OUTPUT
    flowSP : REAL;
    valveCommand : REAL;
    fault : BOOL;
    normalMode : BOOL;
END_VAR
VAR
    initDone : BOOL := FALSE;
    prevMode : INT := 0;
    prevReset : BOOL := FALSE;
    prevFlowSP : REAL := 0.0;
    prevValveCommand : REAL := 0.0;
    accT : REAL := 0.0;
    accF : REAL := 0.0;
    tempError : REAL;
    flowError : REAL;
    trialT : REAL;
    trialF : REAL;
    rawFlow : REAL;
    rawValve : REAL;
    modeChanged : BOOL;
    resetRise : BOOL;
END_VAR

fault := (mode < 0) OR (mode > 2) OR (scanSeconds <= 0.0) OR (scanSeconds > 10.0);
resetRise := resetBtn AND NOT prevReset;
normalMode := FALSE;

IF NOT initDone THEN
    flowSP := manualFlowSP;
    valveCommand := manualValve;
    tempError := tempSP - tempPV;
    accT := flowSP - 1.0 * tempError;
    flowError := flowSP - flowPV;
    accF := valveCommand - 2.0 * flowError;
ELSE
    modeChanged := mode <> prevMode;

    IF resetRise THEN
        flowSP := manualFlowSP;
        valveCommand := manualValve;
        tempError := tempSP - tempPV;
        accT := flowSP - 1.0 * tempError;
        flowError := flowSP - flowPV;
        accF := valveCommand - 2.0 * flowError;
    ELSIF fault THEN
        flowSP := manualFlowSP;
        valveCommand := manualValve;
        tempError := tempSP - tempPV;
        accT := flowSP - 1.0 * tempError;
        flowError := flowSP - flowPV;
        accF := valveCommand - 2.0 * flowError;
    ELSIF modeChanged THEN
        IF mode = 2 THEN
            flowSP := prevFlowSP;
            valveCommand := prevValveCommand;
            tempError := tempSP - tempPV;
            accT := flowSP - 1.0 * tempError;
            flowError := flowSP - flowPV;
            accF := valveCommand - 2.0 * flowError;
        ELSE
            flowSP := manualFlowSP;
            valveCommand := prevValveCommand;
            tempError := tempSP - tempPV;
            accT := flowSP - 1.0 * tempError;
            flowError := flowSP - flowPV;
            accF := valveCommand - 2.0 * flowError;
        END_IF
    ELSE
        normalMode := TRUE;
        IF mode = 0 THEN
            flowSP := manualFlowSP;
            valveCommand := manualValve;
            tempError := tempSP - tempPV;
            accT := flowSP - 1.0 * tempError;
            flowError := flowSP - flowPV;
            accF := valveCommand - 2.0 * flowError;
        ELSIF mode = 1 THEN
            flowSP := manualFlowSP;
            flowError := flowSP - flowPV;
            trialF := accF + 0.5 * flowError * scanSeconds;
            rawValve := 2.0 * flowError + trialF;
            IF rawValve < 0.0 THEN
                valveCommand := 0.0;
            ELSIF rawValve > 100.0 THEN
                valveCommand := 100.0;
            ELSE
                valveCommand := rawValve;
            END_IF
            accF := valveCommand - 2.0 * flowError;
            tempError := tempSP - tempPV;
            accT := flowSP - 1.0 * tempError;
        ELSE
            tempError := tempSP - tempPV;
            trialT := accT + 0.2 * tempError * scanSeconds;
            rawFlow := 1.0 * tempError + trialT;
            IF rawFlow < 0.0 THEN
                flowSP := 0.0;
            ELSIF rawFlow > 50.0 THEN
                flowSP := 50.0;
            ELSE
                flowSP := rawFlow;
            END_IF
            accT := flowSP - 1.0 * tempError;

            flowError := flowSP - flowPV;
            trialF := accF + 0.5 * flowError * scanSeconds;
            rawValve := 2.0 * flowError + trialF;
            IF rawValve < 0.0 THEN
                valveCommand := 0.0;
            ELSIF rawValve > 100.0 THEN
                valveCommand := 100.0;
            ELSE
                valveCommand := rawValve;
            END_IF
            accF := valveCommand - 2.0 * flowError;
        END_IF
    END_IF
END_IF

prevMode := mode;
prevReset := resetBtn;
prevFlowSP := flowSP;
prevValveCommand := valveCommand;
initDone := TRUE;
END_FUNCTION_BLOCK

(* ---- self-medium-01.candidate_01.st ---- *)
TYPE ST_Recipe :
STRUCT
    recipeID : INT;
    totalRatio : REAL;
    temperature : REAL;
END_STRUCT;
END_TYPE;

FUNCTION_BLOCK FB
VAR_INPUT
    recipe : ARRAY[1..8] OF ST_Recipe;
    selSlot : INT;
    loadCmd : BOOL;
    running : BOOL;
END_VAR
VAR_OUTPUT
    valid : BOOL;
    loadedID : INT;
END_VAR
VAR
    loadCmdPrevious : BOOL;
    loadEdge : BOOL;
    slotInRange : BOOL;
    ratioInRange : BOOL;
    tempInRange : BOOL;
    slotOccupied : BOOL;
    latchedValid : BOOL;
    latchedLoadedID : INT;
END_VAR

loadEdge := loadCmd AND NOT loadCmdPrevious;

IF loadEdge AND NOT running THEN
    slotInRange := (selSlot >= 1) AND (selSlot <= 8);

    IF slotInRange THEN
        slotOccupied := (recipe[selSlot].recipeID <> 0);
        ratioInRange := (recipe[selSlot].totalRatio >= 99.0) AND
                        (recipe[selSlot].totalRatio <= 101.0);
        tempInRange := (recipe[selSlot].temperature >= 30.0) AND
                       (recipe[selSlot].temperature <= 180.0);

        latchedValid := slotOccupied AND ratioInRange AND tempInRange;

        IF latchedValid THEN
            latchedLoadedID := recipe[selSlot].recipeID;
        ELSE
            latchedLoadedID := 0;
        END_IF;
    ELSE
        latchedValid := FALSE;
        latchedLoadedID := 0;
    END_IF;
END_IF;

valid := latchedValid;
loadedID := latchedLoadedID;
loadCmdPrevious := loadCmd;

END_FUNCTION_BLOCK

(* ---- self-medium-01.candidate_02.st ---- *)
TYPE ST_Recipe :
STRUCT
    recipeID : INT;
    totalRatio : REAL;
    temperature : REAL;
END_STRUCT;
END_TYPE;

FUNCTION_BLOCK FB
VAR_INPUT
    recipe : ARRAY[1..8] OF ST_Recipe;
    selSlot : INT;
    loadCmd : BOOL;
    running : BOOL;
END_VAR
VAR_OUTPUT
    valid : BOOL;
    loadedID : INT;
END_VAR
VAR
    loadCmdPrevious : BOOL;
    loadEdge : BOOL;
    slotInRange : BOOL;
    ratioInRange : BOOL;
    tempInRange : BOOL;
    slotOccupied : BOOL;
    latchedValid : BOOL;
    latchedLoadedID : INT;
END_VAR

loadEdge := loadCmd AND NOT loadCmdPrevious;

IF loadEdge AND NOT running THEN
    slotInRange := (selSlot >= 1) AND (selSlot <= 8);

    IF slotInRange THEN
        slotOccupied := (recipe[selSlot].recipeID <> 0);
        ratioInRange := (recipe[selSlot].totalRatio >= 99.0) AND
                        (recipe[selSlot].totalRatio <= 101.0);
        tempInRange := (recipe[selSlot].temperature >= 30.0) AND
                       (recipe[selSlot].temperature <= 180.0);

        latchedValid := slotOccupied AND ratioInRange AND tempInRange;

        IF latchedValid THEN
            latchedLoadedID := recipe[selSlot].recipeID;
        ELSE
            latchedLoadedID := 0;
        END_IF;
    ELSE
        latchedValid := FALSE;
        latchedLoadedID := 0;
    END_IF;
END_IF;

valid := latchedValid;
loadedID := latchedLoadedID;
loadCmdPrevious := loadCmd;

END_FUNCTION_BLOCK

(* ---- self-medium-01.raw_candidate_01.st ---- *)
TYPE ST_Recipe :
STRUCT
    recipeID : INT;
    totalRatio : REAL;
    temperature : REAL;
END_STRUCT
END_TYPE

FUNCTION_BLOCK FB
VAR_INPUT
    recipe : ARRAY[1..8] OF ST_Recipe;
    selSlot : INT;
    loadCmd : BOOL;
    running : BOOL;
END_VAR
VAR_OUTPUT
    valid : BOOL;
    loadedID : INT;
END_VAR
VAR
    loadCmdPrevious : BOOL;
    loadEdge : BOOL;
    slotInRange : BOOL;
    ratioInRange : BOOL;
    tempInRange : BOOL;
    slotOccupied : BOOL;
    latchedValid : BOOL;
    latchedLoadedID : INT;
END_VAR

loadEdge := loadCmd AND NOT loadCmdPrevious;

IF loadEdge AND NOT running THEN
    slotInRange := (selSlot >= 1) AND (selSlot <= 8);

    IF slotInRange THEN
        slotOccupied := (recipe[selSlot].recipeID <> 0);
        ratioInRange := (recipe[selSlot].totalRatio >= 99.0) AND
                        (recipe[selSlot].totalRatio <= 101.0);
        tempInRange := (recipe[selSlot].temperature >= 30.0) AND
                       (recipe[selSlot].temperature <= 180.0);

        latchedValid := slotOccupied AND ratioInRange AND tempInRange;

        IF latchedValid THEN
            latchedLoadedID := recipe[selSlot].recipeID;
        ELSE
            latchedLoadedID := 0;
        END_IF;
    ELSE
        latchedValid := FALSE;
        latchedLoadedID := 0;
    END_IF;
END_IF;

valid := latchedValid;
loadedID := latchedLoadedID;
loadCmdPrevious := loadCmd;

END_FUNCTION_BLOCK

(* ---- self-medium-01.raw_candidate_02.st ---- *)
TYPE ST_Recipe :
STRUCT
    recipeID : INT;
    totalRatio : REAL;
    temperature : REAL;
END_STRUCT
END_TYPE

FUNCTION_BLOCK FB
VAR_INPUT
    recipe : ARRAY[1..8] OF ST_Recipe;
    selSlot : INT;
    loadCmd : BOOL;
    running : BOOL;
END_VAR
VAR_OUTPUT
    valid : BOOL;
    loadedID : INT;
END_VAR
VAR
    loadCmdPrevious : BOOL;
    loadEdge : BOOL;
    slotInRange : BOOL;
    ratioInRange : BOOL;
    tempInRange : BOOL;
    slotOccupied : BOOL;
    latchedValid : BOOL;
    latchedLoadedID : INT;
END_VAR

loadEdge := loadCmd AND NOT loadCmdPrevious;

IF loadEdge AND NOT running THEN
    slotInRange := (selSlot >= 1) AND (selSlot <= 8);

    IF slotInRange THEN
        slotOccupied := (recipe[selSlot].recipeID <> 0);
        ratioInRange := (recipe[selSlot].totalRatio >= 99.0) AND
                        (recipe[selSlot].totalRatio <= 101.0);
        tempInRange := (recipe[selSlot].temperature >= 30.0) AND
                       (recipe[selSlot].temperature <= 180.0);

        latchedValid := slotOccupied AND ratioInRange AND tempInRange;

        IF latchedValid THEN
            latchedLoadedID := recipe[selSlot].recipeID;
        ELSE
            latchedLoadedID := 0;
        END_IF;
    ELSE
        latchedValid := FALSE;
        latchedLoadedID := 0;
    END_IF;
END_IF;

valid := latchedValid;
loadedID := latchedLoadedID;
loadCmdPrevious := loadCmd;

END_FUNCTION_BLOCK

(* ---- self-medium-02.candidate_01.st ---- *)
FUNCTION_BLOCK FB
VAR_INPUT
    enable : BOOL;
    rawValue : REAL;
END_VAR
VAR_OUTPUT
    filteredValue : REAL;
    windowFull : BOOL;
    sampleCount : INT;
END_VAR
VAR
    buffer : ARRAY[0..7] OF REAL;
    writeIndex : INT;
    bufIdx : INT;
    sum : REAL;
END_VAR

IF NOT enable THEN
    sampleCount := 0;
    windowFull := FALSE;
    writeIndex := 0;
    FOR bufIdx := 0 TO 7 DO
        buffer[bufIdx] := 0.0;
    END_FOR;
ELSE
    buffer[writeIndex] := rawValue;

    writeIndex := writeIndex + 1;
    IF writeIndex >= 8 THEN
        writeIndex := 0;
    END_IF;

    IF sampleCount < 8 THEN
        sampleCount := sampleCount + 1;
    END_IF;

    sum := 0.0;
    FOR bufIdx := 0 TO sampleCount - 1 DO
        sum := sum + buffer[bufIdx];
    END_FOR;

    filteredValue := sum / INT_TO_REAL(sampleCount);
    windowFull := sampleCount >= 8;
END_IF;

END_FUNCTION_BLOCK

(* ---- self-medium-02.raw_candidate_01.st ---- *)
FUNCTION_BLOCK FB
VAR_INPUT
    enable : BOOL;
    rawValue : REAL;
END_VAR
VAR_OUTPUT
    filteredValue : REAL;
    windowFull : BOOL;
    sampleCount : INT;
END_VAR
VAR
    buffer : ARRAY[0..7] OF REAL;
    writeIndex : INT;
    bufIdx : INT;
    sum : REAL;
END_VAR

IF NOT enable THEN
    sampleCount := 0;
    windowFull := FALSE;
    writeIndex := 0;
    FOR bufIdx := 0 TO 7 DO
        buffer[bufIdx] := 0.0;
    END_FOR;
ELSE
    buffer[writeIndex] := rawValue;

    writeIndex := writeIndex + 1;
    IF writeIndex >= 8 THEN
        writeIndex := 0;
    END_IF;

    IF sampleCount < 8 THEN
        sampleCount := sampleCount + 1;
    END_IF;

    sum := 0.0;
    FOR bufIdx := 0 TO sampleCount - 1 DO
        sum := sum + buffer[bufIdx];
    END_FOR;

    filteredValue := sum / INT_TO_REAL(sampleCount);
    windowFull := sampleCount >= 8;
END_IF;

END_FUNCTION_BLOCK

(* ---- self-medium-03.candidate_01.st ---- *)
FUNCTION_BLOCK FB
VAR_INPUT
    openBtn: BOOL;
    closeBtn: BOOL;
    openLimit: BOOL;
    closeLimit: BOOL;
    obstacle: BOOL;
END_VAR
VAR_OUTPUT
    motorUp: BOOL;
    motorDown: BOOL;
    errorFlag: BOOL;
END_VAR
VAR
    prevOpenBtn: BOOL := FALSE;
    prevCloseBtn: BOOL := FALSE;
    prevMotorUp: BOOL := FALSE;
    prevMotorDown: BOOL := FALSE;
    prevErrorFlag: BOOL := FALSE;
    openRising: BOOL;
    closeRising: BOOL;
    bothRising: BOOL;
END_VAR

openRising := openBtn AND (NOT prevOpenBtn);
closeRising := closeBtn AND (NOT prevCloseBtn);
bothRising := (openBtn AND closeBtn) AND (NOT (prevOpenBtn AND prevCloseBtn));

motorUp := (NOT obstacle) AND (NOT openLimit) AND
    (prevMotorUp OR
     ((NOT prevMotorUp) AND (NOT prevMotorDown) AND (NOT prevErrorFlag) AND
      openRising AND (NOT closeBtn)));

motorDown := (NOT obstacle) AND (NOT closeLimit) AND
    (prevMotorDown OR
     ((NOT prevMotorUp) AND (NOT prevMotorDown) AND (NOT prevErrorFlag) AND
      closeRising AND (NOT openBtn)));

errorFlag := obstacle OR (prevErrorFlag AND (NOT bothRising));

prevOpenBtn := openBtn;
prevCloseBtn := closeBtn;
prevMotorUp := motorUp;
prevMotorDown := motorDown;
prevErrorFlag := errorFlag;

END_FUNCTION_BLOCK

(* ---- self-medium-03.raw_candidate_01.st ---- *)
FUNCTION_BLOCK FB
VAR_INPUT
    openBtn: BOOL;
    closeBtn: BOOL;
    openLimit: BOOL;
    closeLimit: BOOL;
    obstacle: BOOL;
END_VAR
VAR_OUTPUT
    motorUp: BOOL;
    motorDown: BOOL;
    errorFlag: BOOL;
END_VAR
VAR
    prevOpenBtn: BOOL := FALSE;
    prevCloseBtn: BOOL := FALSE;
    prevMotorUp: BOOL := FALSE;
    prevMotorDown: BOOL := FALSE;
    prevErrorFlag: BOOL := FALSE;
    openRising: BOOL;
    closeRising: BOOL;
    bothRising: BOOL;
END_VAR

openRising := openBtn AND (NOT prevOpenBtn);
closeRising := closeBtn AND (NOT prevCloseBtn);
bothRising := (openBtn AND closeBtn) AND (NOT (prevOpenBtn AND prevCloseBtn));

motorUp := (NOT obstacle) AND (NOT openLimit) AND
    (prevMotorUp OR
     ((NOT prevMotorUp) AND (NOT prevMotorDown) AND (NOT prevErrorFlag) AND
      openRising AND (NOT closeBtn)));

motorDown := (NOT obstacle) AND (NOT closeLimit) AND
    (prevMotorDown OR
     ((NOT prevMotorUp) AND (NOT prevMotorDown) AND (NOT prevErrorFlag) AND
      closeRising AND (NOT openBtn)));

errorFlag := obstacle OR (prevErrorFlag AND (NOT bothRising));

prevOpenBtn := openBtn;
prevCloseBtn := closeBtn;
prevMotorUp := motorUp;
prevMotorDown := motorDown;
prevErrorFlag := errorFlag;

END_FUNCTION_BLOCK

(* ---- self-medium-04.candidate_01.st ---- *)
FUNCTION_BLOCK FB
VAR_INPUT
    startBtn : BOOL;
    resetBtn : BOOL;
    doneSensor : BOOL;
    targetVol : REAL;
    flowVol : REAL;
END_VAR
VAR_OUTPUT
    valveOpen : BOOL;
    fillsToday : INT;
END_VAR
VAR
    prevStartBtn : BOOL := FALSE;
    prevResetBtn : BOOL := FALSE;
    prevValveOpen : BOOL := FALSE;
    accumulatedVolume : REAL := 0.0;
    pendingConfirm : BOOL := FALSE;
    startEdge : BOOL;
    resetEdge : BOOL;
    fillingNow : BOOL;
END_VAR

startEdge := startBtn AND NOT prevStartBtn;
resetEdge := resetBtn AND NOT prevResetBtn;

IF resetEdge THEN
    fillsToday := 0;
    accumulatedVolume := 0.0;
    pendingConfirm := FALSE;
    valveOpen := FALSE;
ELSE
    fillingNow := prevValveOpen;

    IF startEdge AND NOT prevValveOpen THEN
        pendingConfirm := FALSE;
        accumulatedVolume := 0.0;
        valveOpen := TRUE;
        fillingNow := TRUE;
    END_IF;

    IF fillingNow THEN
        accumulatedVolume := accumulatedVolume + flowVol;

        IF accumulatedVolume >= targetVol THEN
            valveOpen := FALSE;
            pendingConfirm := TRUE;
        ELSE
            valveOpen := TRUE;
        END_IF;
    END_IF;

    IF pendingConfirm AND doneSensor AND NOT valveOpen THEN
        IF fillsToday < 32767 THEN
            fillsToday := fillsToday + 1;
        END_IF;
        pendingConfirm := FALSE;
    END_IF;
END_IF;

prevStartBtn := startBtn;
prevResetBtn := resetBtn;
prevValveOpen := valveOpen;
END_FUNCTION_BLOCK

(* ---- self-medium-04.raw_candidate_01.st ---- *)
FUNCTION_BLOCK FB
VAR_INPUT
    startBtn : BOOL;
    resetBtn : BOOL;
    doneSensor : BOOL;
    targetVol : REAL;
    flowVol : REAL;
END_VAR
VAR_OUTPUT
    valveOpen : BOOL;
    fillsToday : INT;
END_VAR
VAR
    prevStartBtn : BOOL := FALSE;
    prevResetBtn : BOOL := FALSE;
    prevValveOpen : BOOL := FALSE;
    accumulatedVolume : REAL := 0.0;
    pendingConfirm : BOOL := FALSE;
    startEdge : BOOL;
    resetEdge : BOOL;
    fillingNow : BOOL;
END_VAR

startEdge := startBtn AND NOT prevStartBtn;
resetEdge := resetBtn AND NOT prevResetBtn;

IF resetEdge THEN
    fillsToday := 0;
    accumulatedVolume := 0.0;
    pendingConfirm := FALSE;
    valveOpen := FALSE;
ELSE
    fillingNow := prevValveOpen;

    IF startEdge AND NOT prevValveOpen THEN
        pendingConfirm := FALSE;
        accumulatedVolume := 0.0;
        valveOpen := TRUE;
        fillingNow := TRUE;
    END_IF;

    IF fillingNow THEN
        accumulatedVolume := accumulatedVolume + flowVol;

        IF accumulatedVolume >= targetVol THEN
            valveOpen := FALSE;
            pendingConfirm := TRUE;
        ELSE
            valveOpen := TRUE;
        END_IF;
    END_IF;

    IF pendingConfirm AND doneSensor AND NOT valveOpen THEN
        IF fillsToday < 32767 THEN
            fillsToday := fillsToday + 1;
        END_IF;
        pendingConfirm := FALSE;
    END_IF;
END_IF;

prevStartBtn := startBtn;
prevResetBtn := resetBtn;
prevValveOpen := valveOpen;
END_FUNCTION_BLOCK

(* ---- self-medium-05.candidate_01.st ---- *)
FUNCTION_BLOCK FB
VAR_INPUT
    enable : BOOL;
    resetBtn : BOOL;
    scanSeconds : LREAL;
    steamFlow : LREAL;
    fuelFlow : LREAL;
    steamTemp : LREAL;
    steamPressure : LREAL;
END_VAR
VAR_OUTPUT
    qualified : BOOL;
    dataFault : BOOL;
    qualifiedTon : LREAL;
    fuelTon : LREAL;
    revenue : LREAL;
    cost : LREAL;
    netProfit : LREAL;
END_VAR
VAR
    prevResetBtn : BOOL;
    resetRising : BOOL;
    tonAccQualified : LREAL;
    tonAccFuel : LREAL;
END_VAR

resetRising := resetBtn AND NOT prevResetBtn;

qualified := steamTemp >= 447.0 AND steamTemp <= 453.0 AND steamPressure >= 3750.0 AND steamPressure <= 3850.0;

dataFault := scanSeconds <= 0.0 OR scanSeconds > 10.0 OR steamFlow < 0.0 OR steamFlow > 90.0 OR fuelFlow < 0.0 OR fuelFlow > 6.0;

IF resetRising THEN
    tonAccQualified := 0.0;
    tonAccFuel := 0.0;
ELSIF enable AND NOT dataFault THEN
    tonAccFuel := tonAccFuel + fuelFlow * scanSeconds / 1000.0;
    IF qualified THEN
        tonAccQualified := tonAccQualified + steamFlow * scanSeconds / 1000.0;
    END_IF;
END_IF;

qualifiedTon := tonAccQualified;
fuelTon := tonAccFuel;
revenue := tonAccQualified * 280.0;
cost := tonAccFuel * 1500.0;
netProfit := revenue - cost;

prevResetBtn := resetBtn;

END_FUNCTION_BLOCK

(* ---- self-medium-05.raw_candidate_01.st ---- *)
FUNCTION_BLOCK FB
VAR_INPUT
    enable : BOOL;
    resetBtn : BOOL;
    scanSeconds : LREAL;
    steamFlow : LREAL;
    fuelFlow : LREAL;
    steamTemp : LREAL;
    steamPressure : LREAL;
END_VAR
VAR_OUTPUT
    qualified : BOOL;
    dataFault : BOOL;
    qualifiedTon : LREAL;
    fuelTon : LREAL;
    revenue : LREAL;
    cost : LREAL;
    netProfit : LREAL;
END_VAR
VAR
    prevResetBtn : BOOL;
    resetRising : BOOL;
    tonAccQualified : LREAL;
    tonAccFuel : LREAL;
END_VAR

resetRising := resetBtn AND NOT prevResetBtn;

qualified := steamTemp >= 447.0 AND steamTemp <= 453.0 AND steamPressure >= 3750.0 AND steamPressure <= 3850.0;

dataFault := scanSeconds <= 0.0 OR scanSeconds > 10.0 OR steamFlow < 0.0 OR steamFlow > 90.0 OR fuelFlow < 0.0 OR fuelFlow > 6.0;

IF resetRising THEN
    tonAccQualified := 0.0;
    tonAccFuel := 0.0;
ELSIF enable AND NOT dataFault THEN
    tonAccFuel := tonAccFuel + fuelFlow * scanSeconds / 1000.0;
    IF qualified THEN
        tonAccQualified := tonAccQualified + steamFlow * scanSeconds / 1000.0;
    END_IF
END_IF

qualifiedTon := tonAccQualified;
fuelTon := tonAccFuel;
revenue := tonAccQualified * 280.0;
cost := tonAccFuel * 1500.0;
netProfit := revenue - cost;

prevResetBtn := resetBtn;

END_FUNCTION_BLOCK

(* ---- self-medium-06.candidate_01.st ---- *)
FUNCTION_BLOCK FB
VAR_INPUT
    enable : BOOL;
    resetBtn : BOOL;
    sensorValid : BOOL;
    setpoint : REAL;
    temperature : REAL;
    scanSeconds : REAL;
    bias : REAL;
END_VAR
VAR_OUTPUT
    power : REAL;
    correction : REAL;
    fault : BOOL;
END_VAR
VAR
    ePrev : REAL := 0.0;
    historyValid : BOOL := FALSE;
    resetPrev : BOOL := FALSE;
    resetRising : BOOL;
    e : REAL;
    de : REAL;
    x : REAL;
    y : REAL;
END_VAR

resetRising := resetBtn AND NOT resetPrev;
fault := (NOT sensorValid) OR (scanSeconds <= 0.0) OR (scanSeconds > 10.0);

IF (NOT enable) OR fault OR resetRising THEN
    power := 0.0;
    correction := 0.0;
    ePrev := 0.0;
    historyValid := FALSE;
ELSE
    e := setpoint - temperature;

    IF NOT historyValid THEN
        de := 0.0;
    ELSE
        de := (e - ePrev) / scanSeconds;
    END_IF;

    x := LIMIT(-1.0, e / 10.0, 1.0);
    y := LIMIT(-1.0, de / 2.0, 1.0);

    correction := 20.0 * x + 10.0 * y;
    power := LIMIT(0.0, bias + correction, 100.0);

    ePrev := e;
    historyValid := TRUE;
END_IF;

resetPrev := resetBtn;

END_FUNCTION_BLOCK

(* ---- self-medium-06.raw_candidate_01.st ---- *)
FUNCTION_BLOCK FB
VAR_INPUT
    enable : BOOL;
    resetBtn : BOOL;
    sensorValid : BOOL;
    setpoint : REAL;
    temperature : REAL;
    scanSeconds : REAL;
    bias : REAL;
END_VAR
VAR_OUTPUT
    power : REAL;
    correction : REAL;
    fault : BOOL;
END_VAR
VAR
    ePrev : REAL := 0.0;
    historyValid : BOOL := FALSE;
    resetPrev : BOOL := FALSE;
    resetRising : BOOL;
    e : REAL;
    de : REAL;
    x : REAL;
    y : REAL;
END_VAR

resetRising := resetBtn AND NOT resetPrev;
fault := (NOT sensorValid) OR (scanSeconds <= 0.0) OR (scanSeconds > 10.0);

IF (NOT enable) OR fault OR resetRising THEN
    power := 0.0;
    correction := 0.0;
    ePrev := 0.0;
    historyValid := FALSE;
ELSE
    e := setpoint - temperature;

    IF NOT historyValid THEN
        de := 0.0;
    ELSE
        de := (e - ePrev) / scanSeconds;
    END_IF;

    x := LIMIT(-1.0, e / 10.0, 1.0);
    y := LIMIT(-1.0, de / 2.0, 1.0);

    correction := 20.0 * x + 10.0 * y;
    power := LIMIT(0.0, bias + correction, 100.0);

    ePrev := e;
    historyValid := TRUE;
END_IF;

resetPrev := resetBtn;

END_FUNCTION_BLOCK
